FUNCTION "FRK_UnitRelease" : Void   // FC79, SCL
{ S7_Optimized_Access := 'TRUE' }
VERSION : 0.1
// stored: AutoNumber true, IsIECCheckEnabled false, SetENOAutomatically false, UDAEnableTagReadback false
   VAR_INPUT
      Gate : DInt;
      Desired : DInt;
      Trusted : Bool;
      Core : "FRK_Core";
      Unit : "FRK_Unit";
      Status : "ST_ModuleStatus";
      Policy : Array[0..6] of "ST_ModePolicy";
      Access : "FRK_Access";
      Supported : Array[0..6] of Bool;
   END_VAR
   VAR_IN_OUT
      Report : "ST_ReleaseReport";
   END_VAR
BEGIN

   #Report.Count := 0;
   #Report.Released := TRUE;
   IF #Gate <> 5 AND #Gate <> 4
       AND #Gate <> 7 AND #Gate <> 2
       AND #Gate <> 8
       AND NOT (#Unit.ConfigEnabled AND #Gate = 1)
       AND NOT (#Unit.ConfigSetsEnabled AND #Gate = 11)
       AND NOT (#Unit.ModelEnabled AND #Gate = 3) THEN
       "FRK_ReleaseReason"(Report := #Report,
                           Description := WSTRING#'std.error.unsupportedHmiRequest',
                           Reason := 2008,
                           Path := STRING_TO_WSTRING(#Status.Name),
                           Kind := 4);
       RETURN;
   END_IF;
   IF NOT #Trusted THEN
       IF #Access.CurrentLevel < #Access.Policy.Required[#Gate] THEN
           "FRK_ReleaseReason"(Report := #Report,
                               Description := WSTRING#'std.release.insufficientAction',
                               Reason := 2002,
                               Path := STRING_TO_WSTRING(#Status.Name),
                               Kind := 1);
       END_IF;
   END_IF;
   CASE #Gate OF
       3:
           IF #Core.Exec <> 0 OR #Unit.ModePending OR #Unit.Clearing OR NOT "FRK_DescendantsReady"(OwnerIndex := #Core.RegIndex) THEN
               "FRK_ReleaseReason"(Report := #Report,
                                   Description := WSTRING#'std.error.hmiRequestRejected',
                                   Reason := 2011,
                                   Path := STRING_TO_WSTRING(#Status.Name),
                                   Kind := 4);
           END_IF;
           IF #Unit.AlarmBlocking THEN
               "FRK_ReleaseReason"(Report := #Report,
                                   Description := WSTRING#'std.release.manualReset',
                                   Reason := 0,
                                   Path := STRING_TO_WSTRING(#Status.Name),
                                   Kind := 2);
           END_IF;
           IF NOT #Unit.Permit THEN
               "FRK_ReleaseReason"(Report := #Report,
                                   Description := #Unit.PermitDiag.Description,
                                   Reason := #Unit.PermitDiag.ReasonCode,
                                   Path := #Unit.PermitDiag.SourcePath,
                                   Kind := 3);
           END_IF;
       5:
           // Desired=0 is Start, Desired=1 is Stop. Generic action query is Stop.
           IF #Desired = 0 THEN
               IF #Unit.Mode = 1 OR #Unit.ModePending THEN
                   "FRK_ReleaseReason"(Report := #Report,
                                       Description := WSTRING#'std.error.unsupportedModeRequest',
                                       Reason := 2002,
                                       Path := STRING_TO_WSTRING(#Status.Name),
                                       Kind := 0);
               END_IF;
               IF #Core.Exec <> 0 OR #Unit.RunReq OR #Unit.Clearing OR #Unit.FaultLatched THEN
                   "FRK_ReleaseReason"(Report := #Report,
                                       Description := WSTRING#'std.error.hmiRequestRejected',
                                       Reason := 2011,
                                       Path := STRING_TO_WSTRING(#Status.Name),
                                       Kind := 4);
               END_IF;
               IF #Unit.AlarmBlocking THEN
                   "FRK_ReleaseReason"(Report := #Report,
                                       Description := WSTRING#'std.release.manualReset',
                                       Reason := 0,
                                       Path := STRING_TO_WSTRING(#Status.Name),
                                       Kind := 2);
               END_IF;
               IF #Unit.ConfigBlocked THEN
                   "FRK_ReleaseReason"(Report := #Report,
                                       Description := WSTRING#'std.release.configRestoreUnacknowledged',
                                       Reason := 2040,
                                       Path := STRING_TO_WSTRING(#Status.Name),
                                       Kind := 2);
               END_IF;
               IF NOT #Unit.Permit THEN
                   "FRK_ReleaseReason"(Report := #Report,
                                       Description := #Unit.PermitDiag.Description,
                                       Reason := #Unit.PermitDiag.ReasonCode,
                                       Path := #Unit.PermitDiag.SourcePath,
                                       Kind := 3);
               END_IF;
           END_IF;
       4:
           IF #Unit.ModePending THEN
               "FRK_ReleaseReason"(Report := #Report,
                                   Description := WSTRING#'std.release.modeChangeAlreadyPending',
                                   Reason := 2011,
                                   Path := STRING_TO_WSTRING(#Status.Name),
                                   Kind := 0);
           END_IF;
           IF #Core.Exec = 1 AND #Unit.Mode <> 1 THEN
               IF #Policy[#Unit.Mode].Shield = 2 THEN
                   "FRK_ReleaseReason"(Report := #Report,
                                       Description := WSTRING#'std.release.modeSwitchBlockedWhileRunning',
                                       Reason := 2002,
                                       Path := STRING_TO_WSTRING(#Status.Name),
                                       Kind := 0);
               END_IF;
           END_IF;
           IF #Desired <> -1 THEN
               IF #Desired < 0 OR #Desired >= 7 THEN
                   "FRK_ReleaseReason"(Report := #Report,
                                       Description := WSTRING#'std.error.unsupportedModeRequest',
                                       Reason := 2008,
                                       Path := STRING_TO_WSTRING(#Status.Name),
                                       Kind := 0);
               ELSIF NOT #Supported[#Desired] THEN
                   "FRK_ReleaseReason"(Report := #Report,
                                       Description := WSTRING#'std.error.unsupportedModeRequest',
                                       Reason := 2008,
                                       Path := STRING_TO_WSTRING(#Status.Name),
                                       Kind := 0);
               END_IF;
           END_IF;
       7:
           // The complete alarm model is separate; this gate owns the current latch.
           IF NOT #Unit.FaultLatched AND NOT #Unit.AlarmBlocking AND #Core.Exec = 0 AND NOT #Unit.Clearing AND NOT #Unit.ModePending AND NOT #Unit.FollowStart THEN
               IF "FRK_DescendantsReady"(OwnerIndex := #Core.RegIndex) THEN
                   "FRK_ReleaseReason"(Report := #Report,
                                       Description := WSTRING#'std.release.noBlockingAlarm',
                                       Reason := 2011,
                                       Path := STRING_TO_WSTRING(#Status.Name),
                                       Kind := 4);
               END_IF;
           END_IF;
       2:
           "FRK_ManualCommon"(Core := #Core,
                              Unit := #Unit,
                              Status := #Status,
                              Report := #Report);
       ELSE
           RETURN;
   END_CASE;
END_FUNCTION

FUNCTION "FRK_UnitRunStart" : Void   // FC75, SCL
{ S7_Optimized_Access := 'TRUE' }
VERSION : 0.1
// stored: AutoNumber true, IsIECCheckEnabled false, SetENOAutomatically false, UDAEnableTagReadback false
   VAR_INPUT
      Timeout : Time;
      Label : String;
   END_VAR
   VAR_IN_OUT
      Core : "FRK_Core";
      Status : "ST_ModuleStatus";
   END_VAR
BEGIN

   "FRK_Start"(Core := #Core,
               Status := #Status,
               Supported := TRUE,
               Timeout := #Timeout,
               Label := #Label);
   // A continuous run ends at Stop. Bounded commands/steps own progress timeouts.
   #Core.TimeoutMs := 0;
END_FUNCTION

FUNCTION "FRK_UnitSetLocalCarrier" : Void   // FC62, SCL
{ S7_Optimized_Access := 'TRUE' }
VERSION : 0.1
// stored: AutoNumber true, IsIECCheckEnabled false, SetENOAutomatically false, UDAEnableTagReadback false
   VAR_INPUT
      Index : DInt;
   END_VAR
   VAR_IN_OUT
      Unit : "FRK_Unit";
   END_VAR
BEGIN

   #Unit.CarrierIndex := 0;
   IF #Index < 1 OR #Index > 4 THEN
       RETURN;
   END_IF;
   "FRK_Carriers".Slots[#Index].Enabled := TRUE;
   "FRK_Carriers".Slots[#Index].Kind := 2;
   #Unit.CarrierIndex := #Index;
END_FUNCTION

FUNCTION "FRK_UnitSetPermit" : Void   // FC68, SCL
{ S7_Optimized_Access := 'TRUE' }
VERSION : 0.1
// stored: AutoNumber true, IsIECCheckEnabled false, SetENOAutomatically false, UDAEnableTagReadback false
   VAR_INPUT
      Ok : Bool;
      Diag : "ST_Diagnostic";
   END_VAR
   VAR_IN_OUT
      Unit : "FRK_Unit";
   END_VAR
BEGIN

   #Unit.Permit := #Ok;
   #Unit.PermitDiag := #Diag;
END_FUNCTION

FUNCTION "F_CylinderForcePermit" : Void   // FC158, SCL
{ S7_Optimized_Access := 'TRUE' }
VERSION : 0.1
// stored: AutoNumber true, IsIECCheckEnabled false, SetENOAutomatically false, UDAEnableTagReadback false
   VAR_INPUT
      Permit : Bool;
   END_VAR
   VAR_IN_OUT
      Target : "FB_CylinderCM";
   END_VAR
BEGIN

   // The CM applies its own live extension permit as well, even after Done.
   #Target.Device.Withdrawn := NOT #Permit;
END_FUNCTION

FUNCTION "F_CylinderRelease" : Void   // FC157, SCL
{ S7_Optimized_Access := 'TRUE' }
VERSION : 0.1
// stored: AutoNumber true, IsIECCheckEnabled false, SetENOAutomatically false, UDAEnableTagReadback false
   VAR_IN_OUT
      Seq : "FRK_SequenceCtx";
      Target : "FB_CylinderCM";
   END_VAR
BEGIN

   IF #Target.Device.Lease.Raised AND #Target.Device.Lease.OwnerIndex = #Seq.OwnerIndex
       AND #Target.Device.Lease.ChainIndex = #Seq.ChainIndex AND #Target.Device.Lease.BranchIndex = #Seq.BranchIndex THEN
       #Target.Abort := #Target.Busy;
       #Target.Device.Lease.AbortIssued := #Target.Busy;
       #Target.Execute := FALSE;
       #Target.Device.Lease.Raised := FALSE;
       #Target.Device.Lease.ReleasedScan := #Seq.Scan;
   END_IF;
END_FUNCTION

FUNCTION "F_PressDemoReadInputs" : Void   // FC181, SCL
{ S7_Optimized_Access := 'TRUE' }
VERSION : 0.1
// stored: AutoNumber true, IsIECCheckEnabled false, SetENOAutomatically false, UDAEnableTagReadback false
BEGIN

   "GDB_PressDemoHardwareDriver"(ReadInputs := TRUE);
END_FUNCTION

FUNCTION "F_PressDemoWriteOutputs" : Void   // FC182, SCL
{ S7_Optimized_Access := 'TRUE' }
VERSION : 0.1
// stored: AutoNumber true, IsIECCheckEnabled false, SetENOAutomatically false, UDAEnableTagReadback false
BEGIN

   "GDB_PressDemoHardwareDriver"(ReadInputs := FALSE);
END_FUNCTION

DATA_BLOCK "GDB_FraktalMain"   // DB18
VERSION : 0.1
// stored: AutoNumber true, DBAccessibleFromOPCUA true, DBAccessibleFromWebserver true, InstanceOfName FB_FraktalMain, InstanceOfType FB
"FB_FraktalMain"
BEGIN
END_DATA_BLOCK

DATA_BLOCK "GDB_GRAPH_PressDemoAuto"   // DB14
VERSION : 0.1
// stored: AutoNumber true, DBAccessibleFromOPCUA true, DBAccessibleFromWebserver true, InstanceOfName FB_GRAPH_PressDemoAuto, InstanceOfType FB
"FB_GRAPH_PressDemoAuto"
BEGIN
END_DATA_BLOCK

DATA_BLOCK "GDB_GRAPH_PressDemoHome"   // DB15
VERSION : 0.1
// stored: AutoNumber true, DBAccessibleFromOPCUA true, DBAccessibleFromWebserver true, InstanceOfName FB_GRAPH_PressDemoHome, InstanceOfType FB
"FB_GRAPH_PressDemoHome"
BEGIN
END_DATA_BLOCK

DATA_BLOCK "GDB_PressDemoHardwareDriver"   // DB20
VERSION : 0.1
// stored: AutoNumber true, DBAccessibleFromOPCUA true, DBAccessibleFromWebserver true, InstanceOfName FB_PressDemoHardwareDriver, InstanceOfType FB
"FB_PressDemoHardwareDriver"
BEGIN
END_DATA_BLOCK

DATA_BLOCK "PressDemo"   // DB17
VERSION : 0.1
// stored: AutoNumber true, DBAccessibleFromOPCUA true, DBAccessibleFromWebserver true, InstanceOfName FB_PressDemoUnit, InstanceOfType FB
"FB_PressDemoUnit"
BEGIN
END_DATA_BLOCK
